Fanuc KAREL source: KA00048.KL

PROGRAM KA00048
%NOLOCKGROUP
VAR
  SRC: STRING[80]
  DST: ARRAY[2] OF SHORT
BEGIN
  SRC = 'A'
  DST[1] = SRC
END KA00048
